(* IEC 61131-3 sources: plcassist-cli/packages/volt-lsp-iec/test-corpus/CodesysTestProject/Device/Plc Logic/Application/Library Manager/SysMem, 15 files *)

(* ---- SYSMEMALLOCAREA.fun ---- *)
FUNCTION SYSMEMALLOCAREA : POINTER TO BYTE
VAR_INPUT
	SZCOMPONENT : REFERENCE TO STRING;
	USTYPE : WORD;
	UDISIZE : __XWORD;
	PRESULT : POINTER TO RTS_IEC_RESULT;
END_VAR
END_FUNCTION

(* ---- SYSMEMALLOCCODE.fun ---- *)
FUNCTION SYSMEMALLOCCODE : POINTER TO BYTE
VAR_INPUT
	SZCOMPONENT : REFERENCE TO STRING;
	UDISIZE : __XWORD;
	PRESULT : POINTER TO RTS_IEC_RESULT;
END_VAR
END_FUNCTION

(* ---- SYSMEMALLOCDATA.fun ---- *)
FUNCTION SYSMEMALLOCDATA : POINTER TO BYTE
VAR_INPUT
	SZCOMPONENT : REFERENCE TO STRING;
	UDISIZE : __XWORD;
	PRESULT : POINTER TO RTS_IEC_RESULT;
END_VAR
END_FUNCTION

(* ---- SYSMEMCMP.fun ---- *)
FUNCTION SYSMEMCMP : DINT
VAR_INPUT
	PBUFFER1 : POINTER TO BYTE;
	PBUFFER2 : POINTER TO BYTE;
	UDICOUNT : __XWORD;
END_VAR
END_FUNCTION

(* ---- SYSMEMCPY.fun ---- *)
FUNCTION SYSMEMCPY : POINTER TO BYTE
VAR_INPUT
	PDEST : POINTER TO BYTE;
	PSRC : POINTER TO BYTE;
	UDICOUNT : __XWORD;
END_VAR
END_FUNCTION

(* ---- SYSMEMFORCESWAP.fun ---- *)
FUNCTION SYSMEMFORCESWAP : DINT
VAR_INPUT
	PBYBUFFER : POINTER TO BYTE;
	UDISIZE : UDINT;
	UDICOUNT : UDINT;
END_VAR
END_FUNCTION

(* ---- SYSMEMFREEAREA.fun ---- *)
FUNCTION SYSMEMFREEAREA : RTS_IEC_RESULT
VAR_INPUT
	SZCOMPONENT : REFERENCE TO STRING;
	PMEMORY : POINTER TO BYTE;
END_VAR
END_FUNCTION

(* ---- SYSMEMFREECODE.fun ---- *)
FUNCTION SYSMEMFREECODE : RTS_IEC_RESULT
VAR_INPUT
	SZCOMPONENT : REFERENCE TO STRING;
	PMEMORY : POINTER TO BYTE;
END_VAR
END_FUNCTION

(* ---- SYSMEMFREEDATA.fun ---- *)
FUNCTION SYSMEMFREEDATA : RTS_IEC_RESULT
VAR_INPUT
	SZCOMPONENT : REFERENCE TO STRING;
	PMEMORY : POINTER TO BYTE;
END_VAR
END_FUNCTION

(* ---- SYSMEMGETCURRENTHEAPSIZE.fun ---- *)
FUNCTION SYSMEMGETCURRENTHEAPSIZE : __XWORD
VAR_INPUT
	PRESULT : POINTER TO RTS_IEC_RESULT;
END_VAR
END_FUNCTION

(* ---- SYSMEMISVALIDPOINTER.fun ---- *)
FUNCTION SYSMEMISVALIDPOINTER : RTS_IEC_RESULT
VAR_INPUT
	PTR : POINTER TO BYTE;
	UDISIZE : __XWORD;
	BWRITE : BOOL;
END_VAR
END_FUNCTION

(* ---- SYSMEMMOVE.fun ---- *)
FUNCTION SYSMEMMOVE : POINTER TO BYTE
VAR_INPUT
	PDEST : POINTER TO BYTE;
	PSRC : POINTER TO BYTE;
	UDICOUNT : __XWORD;
END_VAR
END_FUNCTION

(* ---- SYSMEMREALLOCDATA.fun ---- *)
FUNCTION SYSMEMREALLOCDATA : POINTER TO BYTE
VAR_INPUT
	SZCOMPONENT : REFERENCE TO STRING;
	PMEMORY : POINTER TO BYTE;
	UDISIZE : __XWORD;
	PRESULT : POINTER TO RTS_IEC_RESULT;
END_VAR
END_FUNCTION

(* ---- SYSMEMSET.fun ---- *)
FUNCTION SYSMEMSET : POINTER TO BYTE
VAR_INPUT
	PDEST : POINTER TO BYTE;
	UDIVALUE : UDINT;
	UDICOUNT : __XWORD;
END_VAR
END_FUNCTION

(* ---- SYSMEMSWAP.fun ---- *)
FUNCTION SYSMEMSWAP : DINT
VAR_INPUT
	PBYBUFFER : POINTER TO BYTE;
	UDISIZE : UDINT;
	UDICOUNT : UDINT;
END_VAR
END_FUNCTION
